// TIA Portal V19 export
VAR_GLOBAL   // PLC tag table "BT"
   DQ_BT_Green AT %Q0.4 : Bool;
   DQ_BT_Orange AT %Q0.5 : Bool;
   DQ_BT_Red AT %Q0.6 : Bool;
   DQ_BT_Buzzer AT %Q0.7 : Bool;
END_VAR
